// TIA Portal V20 export
// export: Created 2026-10-19T18:45:48.6489181Z, ExportSetting None, DisplayName Totally Integrated Automation Portal, DisplayVersion V20 Update 6, DisplayName TIA Portal Openness, DisplayVersion V20 Update 6, DisplayName TIA Portal Version Control Interface, DisplayVersion V20 Update 6, DisplayName SINAMICS Startdrive Advanced, DisplayVersion V20 SP1, DisplayName SINAMICS Startdrive G130, G150, S120, S150, SINAMICS MV, G220, S200, S210, DisplayVersion V20 SP1, DisplayName SINAMICS Startdrive G110M, G120, G120C, G120D, G120P, G115D, DisplayVersion V20 SP1, DisplayName STEP 7 Professional, DisplayVersion V20 Update 6, DisplayName STEP 7 Safety, DisplayVersion V20 Update 2, DisplayName WinCC Basic/Comfort/Advanced, DisplayVersion V20 Update 6, DisplayName WinCC Unified, DisplayVersion V20 Update 6
VAR_GLOBAL   // PLC tag table "IO_Charger Panel_L3"
   "CHARGER L3 - Output Voltage" AT %ID808 : Real;   // Actual Output Voltage
   "CHARGER L3 - Output Current" AT %ID812 : Real;   // Actual Output Current
   "CHARGER L3 - Set Voltage Feedback" AT %ID816 : Real;   // Set Voltage Value
   "CHARGER L3 - Set Current Feedback" AT %ID820 : Real;   // Set Current Value
   "CHARGER L3 - Charging Start" AT %I824.0 : Bool;   // Charging Running Status
   "CHARGER L3 - Set Voltage Output" AT %QD302 : Real;   // Issue Target Voltage
   "CHARGER L3 - Set Current Output" AT %QD306 : Real;   // Issue Target Current
   "CHARGER L3 - Start Charging" AT %Q310.0 : Bool;   // Start Charging Command
   "CHARGER L3 - Stop Charging" AT %Q310.1 : Bool;   // Stop Charging Command
   "CHARGER L3 - Confirm Voltage & Current Setting" AT %Q310.2 : Bool;   // Confirmation Command
END_VAR
